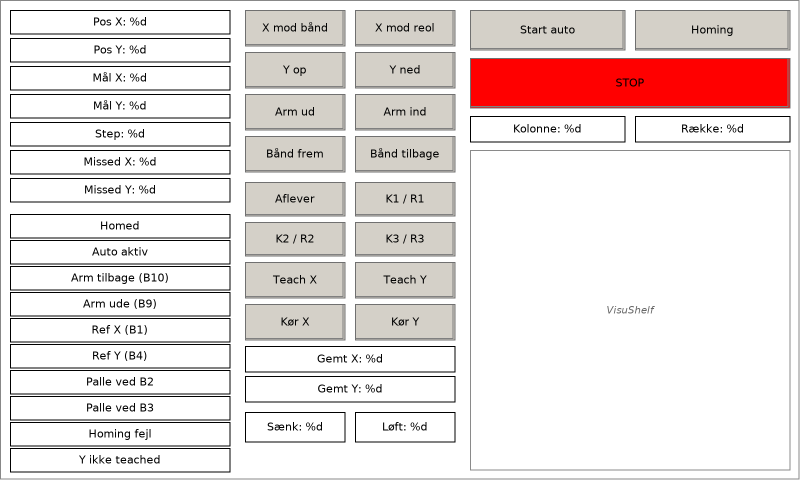
VISUALIZATION VisuTest  // 800x480
    Button (245,10 100x36), "X mod bånd"
        tap MAIN.bJogXBack
    Button (355,10 100x36), "X mod reol"
        tap MAIN.bJogXForward
    Button (245,52 100x36), "Y op"
        tap MAIN.bJogYUp
    Button (355,52 100x36), "Y ned"
        tap MAIN.bJogYDown
    Button (245,94 100x36), "Arm ud"
        tap MAIN.bJogArmOut
    Button (355,94 100x36), "Arm ind"
        tap MAIN.bJogArmIn
    Button (245,136 100x36), "Bånd frem"
        tap MAIN.bJogBeltForward
    Button (355,136 100x36), "Bånd tilbage"
        tap MAIN.bJogBeltBack
    Button (245,262 100x36), "Teach X"
        tap MAIN.bTeachX
    Button (355,262 100x36), "Teach Y"
        tap MAIN.bTeachY
    Button (245,304 100x36), "Kør X"
        tap MAIN.bGoX
    Button (355,304 100x36), "Kør Y"
        tap MAIN.bGoY
    Button (470,10 155x40), "Start auto"
        tap MAIN.bStartAuto
    Button (635,10 155x40), "Homing"
        tap MAIN.bStartHoming
    Button (470,58 320x50), "STOP"
        tap MAIN.bStop
    Rectangle (10,10 220x24), "Pos X: %d", text variable: MAIN.nPosX
    Rectangle (10,38 220x24), "Pos Y: %d", text variable: MAIN.nPosY
    Rectangle (10,66 220x24), "Mål X: %d", text variable: MAIN.nTargetX
    Rectangle (10,94 220x24), "Mål Y: %d", text variable: MAIN.nTargetY
    Rectangle (10,122 220x24), "Step: %d", text variable: MAIN.nStep
    Rectangle (10,150 220x24), "Missed X: %d", text variable: MAIN.nErrorCountX
    Rectangle (10,178 220x24), "Missed Y: %d", text variable: MAIN.nErrorCountY
    Rectangle (245,346 210x26), "Gemt X: %d", text variable: MAIN.nShowX
    Rectangle (245,376 210x26), "Gemt Y: %d", text variable: MAIN.nShowY
    Rectangle (245,412 100x30), "Sænk: %d", text variable: MAIN.nLowerOffset
        OnMouseClick: write the text variable via Default, min 0, max 200
    Rectangle (355,412 100x30), "Løft: %d", text variable: MAIN.nLiftOffset
        OnMouseClick: write the text variable via Default, min 0, max 200
    Rectangle (470,116 155x26), "Kolonne: %d", text variable: MAIN.nSelColumn
    Rectangle (635,116 155x26), "Række: %d", text variable: MAIN.nSelRow
    Rectangle (10,214 220x24), "Homed", colour toggle: MAIN.bHomed
    Rectangle (10,240 220x24), "Auto aktiv", colour toggle: MAIN.bAuto
    Rectangle (10,266 220x24), "Arm tilbage (B10)", colour toggle: MAIN.B10
    Rectangle (10,292 220x24), "Arm ude (B9)", colour toggle: MAIN.B9
    Rectangle (10,318 220x24), "Ref X (B1)", colour toggle: MAIN.B1
    Rectangle (10,344 220x24), "Ref Y (B4)", colour toggle: MAIN.B4
    Rectangle (10,370 220x24), "Palle ved B2", colour toggle: MAIN.bPalletAtB2
    Rectangle (10,396 220x24), "Palle ved B3", colour toggle: MAIN.bPalletAtB3
    Rectangle (10,422 220x24), "Homing fejl", colour toggle: MAIN.bHomingError
    Rectangle (10,448 220x24), "Y ikke teached", colour toggle: MAIN.bYNotTaught
    Frame (470,150 320x320), invisible if: MAIN.bHideShelfSelect
        shows VisuShelf()
    Button (245,182 100x34), "Aflever", colour toggle: MAIN.bSlot0Sel
        OnMouseClick: execute { MAIN.nTeachSlot := 0; }
    Button (355,182 100x34), "K1 / R1", colour toggle: MAIN.bSlot1Sel
        OnMouseClick: execute { MAIN.nTeachSlot := 1; }
    Button (245,222 100x34), "K2 / R2", colour toggle: MAIN.bSlot2Sel
        OnMouseClick: execute { MAIN.nTeachSlot := 2; }
    Button (355,222 100x34), "K3 / R3", colour toggle: MAIN.bSlot3Sel
        OnMouseClick: execute { MAIN.nTeachSlot := 3; }
END_VISUALIZATION

(* stored: Version 1.1.0.1, ProductVersion 3.1.4024.12
   Visu VisuTest: Id {6e3f99c2-464f-4e1a-aa55-836022e67384} *)
